(* IEC 61131-3 sources: llm-plc-st-eval/data/processed_v2/claude-sonnet-4-6/I5/few_shot, 3 files *)

(* ---- ejec_1.st ---- *)
FUNCTION_BLOCK FB_Clasificadora
VAR_INPUT
    sensorPresencia : BOOL; (* Sensor de paso de pieza *)
    sensorAltura    : BOOL; (* Sensor de pieza alta *)
END_VAR
VAR_OUTPUT
    banda   : BOOL; (* Banda transportadora activa *)
    piston  : BOOL; (* Piston desviador *)
    nAltas  : INT;  (* Contador de piezas altas *)
    nBajas  : INT;  (* Contador de piezas bajas *)
END_VAR
VAR
    tRetardo : TON; (* Temporizador de retardo 2 s hasta el desviador *)
    tPulso   : TP;  (* Temporizador de pulso 1 s del piston *)
    rPresencia : R_TRIG; (* Flanco ascendente del sensor de presencia *)
    piezaAlta  : BOOL;   (* Indica que la pieza detectada es alta *)
END_VAR

(* La banda funciona siempre *)
banda := TRUE;

(* Detectar flanco ascendente del sensor de presencia *)
rPresencia(CLK := sensorPresencia);

IF rPresencia.Q THEN
    IF sensorAltura THEN
        (* Pieza alta: registrar y armar retardo *)
        nAltas    := nAltas + 1;
        piezaAlta := TRUE;
    ELSE
        (* Pieza baja: solo contar *)
        nBajas := nBajas + 1;
    END_IF;
END_IF;

(* Retardo de 2 s: la pieza tarda ese tiempo en llegar al desviador *)
tRetardo(IN := piezaAlta, PT := T#2S);

(* Al cumplirse el retardo, lanzar pulso de 1 s en el piston *)
tPulso(IN := tRetardo.Q, PT := T#1S);

(* Activar piston durante el pulso *)
piston := tPulso.Q;

(* Una vez que el pulso termina, liberar el retardo y la bandera *)
IF tPulso.Q = FALSE AND tRetardo.Q = TRUE THEN
    piezaAlta := FALSE;
END_IF;

END_FUNCTION_BLOCK

(* ---- ejec_2.st ---- *)
FUNCTION_BLOCK FB_Clasificadora
VAR_INPUT
    sensorPresencia : BOOL; (* Sensor de paso de pieza *)
    sensorAltura    : BOOL; (* TRUE = pieza alta *)
END_VAR
VAR_OUTPUT
    banda   : BOOL; (* Banda transportadora activa *)
    piston  : BOOL; (* Pistón desviador *)
    nAltas  : INT;  (* Contador de piezas altas *)
    nBajas  : INT;  (* Contador de piezas bajas *)
END_VAR
VAR
    tRetardo : TON; (* Retardo 2 s hasta que la pieza llega al desviador *)
    tPulso   : TP;  (* Pulso 1 s de activación del pistón *)
    rPresencia : R_TRIG; (* Flanco ascendente del sensor de presencia *)
    piezaAlta  : BOOL;   (* Indica que la pieza detectada es alta *)
END_VAR

(* La banda funciona siempre *)
banda := TRUE;

(* Detectar flanco ascendente del sensor de presencia *)
rPresencia(CLK := sensorPresencia);

IF rPresencia.Q THEN
    IF sensorAltura THEN
        (* Pieza alta: registrar y armar retardo *)
        nAltas    := nAltas + 1;
        piezaAlta := TRUE;
    ELSE
        (* Pieza baja: solo contar *)
        nBajas := nBajas + 1;
    END_IF;
END_IF;

(* Retardo de 2 s: empieza cuando se detecta una pieza alta *)
tRetardo(IN := piezaAlta, PT := T#2S);

(* Al cumplirse el retardo, lanzar pulso de 1 s en el pistón *)
tPulso(IN := tRetardo.Q, PT := T#1S);

(* Cuando el pulso termina, limpiar la bandera de pieza alta *)
IF tPulso.Q = FALSE AND tRetardo.Q THEN
    (* El pulso aún no ha terminado; esperar *)
    ;
END_IF;
IF NOT tPulso.Q AND NOT tRetardo.IN THEN
    (* tRetardo.IN vuelve a FALSE solo si piezaAlta = FALSE,
       así que limpiamos piezaAlta cuando el pulso concluye *)
    ;
END_IF;

(* Limpiar piezaAlta una vez que el pulso de 1 s ha finalizado *)
IF tPulso.Q = FALSE AND tRetardo.Q = FALSE AND piezaAlta THEN
    (* El temporizador de retardo ya terminó su ciclo completo *)
    piezaAlta := FALSE;
END_IF;

(* Salida del pistón activa durante el pulso de 1 s *)
piston := tPulso.Q;

END_FUNCTION_BLOCK

(* ---- ejec_3.st ---- *)
FUNCTION_BLOCK FB_Clasificadora
VAR_INPUT
    sensorPresencia : BOOL; (* Sensor de paso de pieza *)
    sensorAltura    : BOOL; (* TRUE = pieza alta *)
END_VAR
VAR_OUTPUT
    banda   : BOOL; (* Banda transportadora activa *)
    piston  : BOOL; (* Pistón desviador *)
    nAltas  : INT;  (* Contador de piezas altas *)
    nBajas  : INT;  (* Contador de piezas bajas *)
END_VAR
VAR
    tRetardo : TON; (* Retardo de 2 s hasta el desviador *)
    tPulso   : TP;  (* Pulso de 1 s para el pistón *)
    rPresencia : R_TRIG; (* Flanco ascendente del sensor de presencia *)
    piezaAlta  : BOOL;   (* Indica que la pieza detectada es alta *)
END_VAR

(* La banda funciona siempre *)
banda := TRUE;

(* Detectar flanco ascendente del sensor de presencia *)
rPresencia(CLK := sensorPresencia);

IF rPresencia.Q THEN
    IF sensorAltura THEN
        (* Pieza alta: registrar y armar retardo *)
        nAltas    := nAltas + 1;
        piezaAlta := TRUE;
    ELSE
        (* Pieza baja: solo contar *)
        nBajas := nBajas + 1;
    END_IF;
END_IF;

(* Retardo de 2 s: comienza cuando hay pieza alta pendiente *)
tRetardo(IN := piezaAlta, PT := T#2S);

(* Al cumplirse el retardo, lanzar pulso de 1 s y limpiar bandera *)
IF tRetardo.Q THEN
    piezaAlta := FALSE; (* Limpiar antes de bajar IN del TON *)
END_IF;

(* Pulso de 1 s para el pistón, disparado por el flanco de tRetardo.Q *)
tPulso(IN := tRetardo.Q, PT := T#1S);

piston := tPulso.Q;

END_FUNCTION_BLOCK
